{attribute 'qualified_only'}
VAR_GLOBAL
	HelloWorld	: STRING;
END_VAR

(* stored: Version 1.1.0.1, ProductVersion 3.1.4024.13
   GVL GVL_Test: Id {aae2f381-adff-43fb-8876-b19caba98a84} *)
